// CFC twin of T_SafeConnection_Tests: the same tests drawn as CFC diagrams, the way a TwinSAFE project is authored.
    FUNCTION_BLOCK T_SafeConnection_Tests_CFC EXTENDS T_SafeCfcTestSuite
    VAR
    // Test_StartsUpToDataWhenGroupRuns
    group_1 : T_SafeGroup;
    conn_1 : T_SafeConnection(group := group_1);
    // Test_ComErrorClearedByAcknowledge
    group_2 : T_SafeGroup;
    conn_2 : T_SafeConnection(group := group_2);
END_VAR

Test_StartsUpToDataWhenGroupRuns();
Test_ComErrorClearedByAcknowledge();

METHOD PRIVATE Test_StartsUpToDataWhenGroupRuns
// note: this text did not pass the execution check against the stored diagram
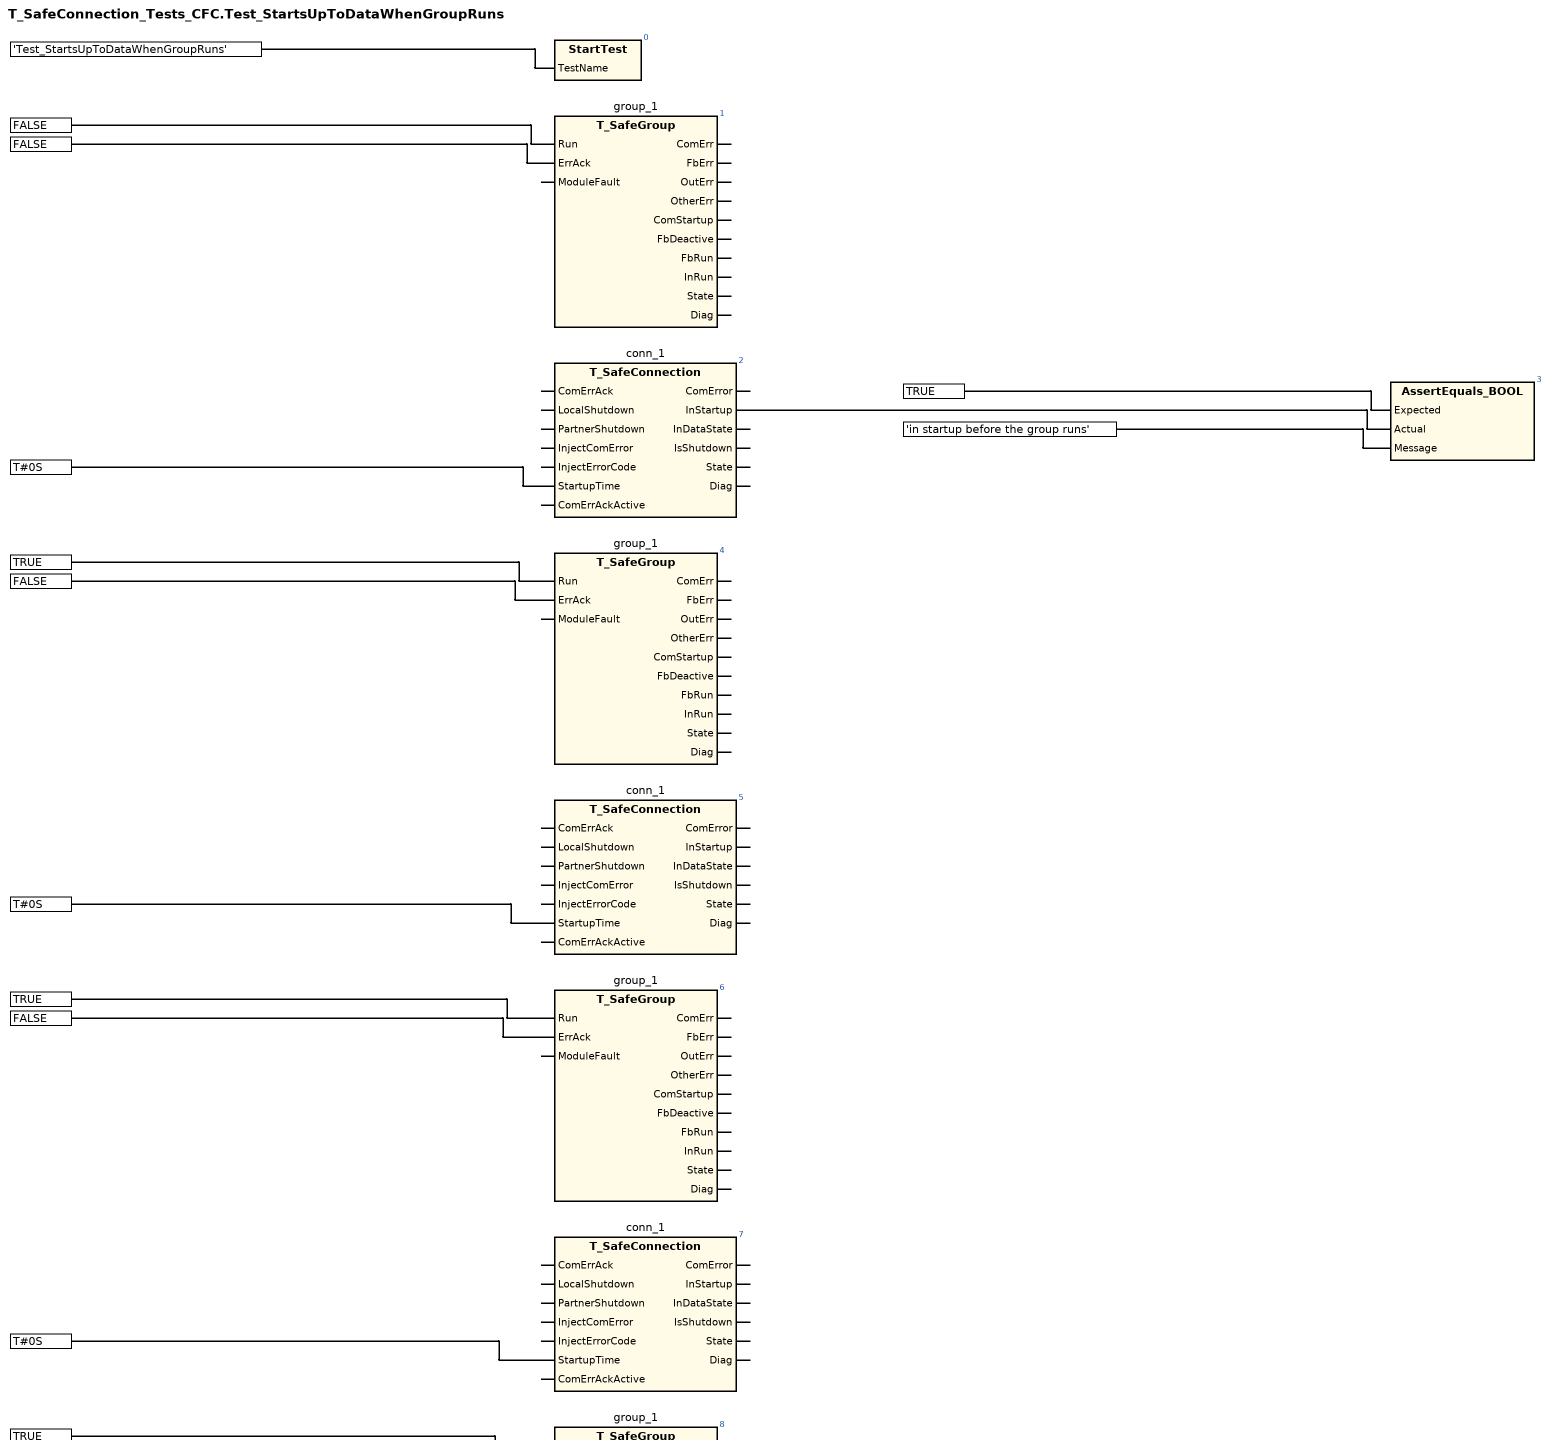
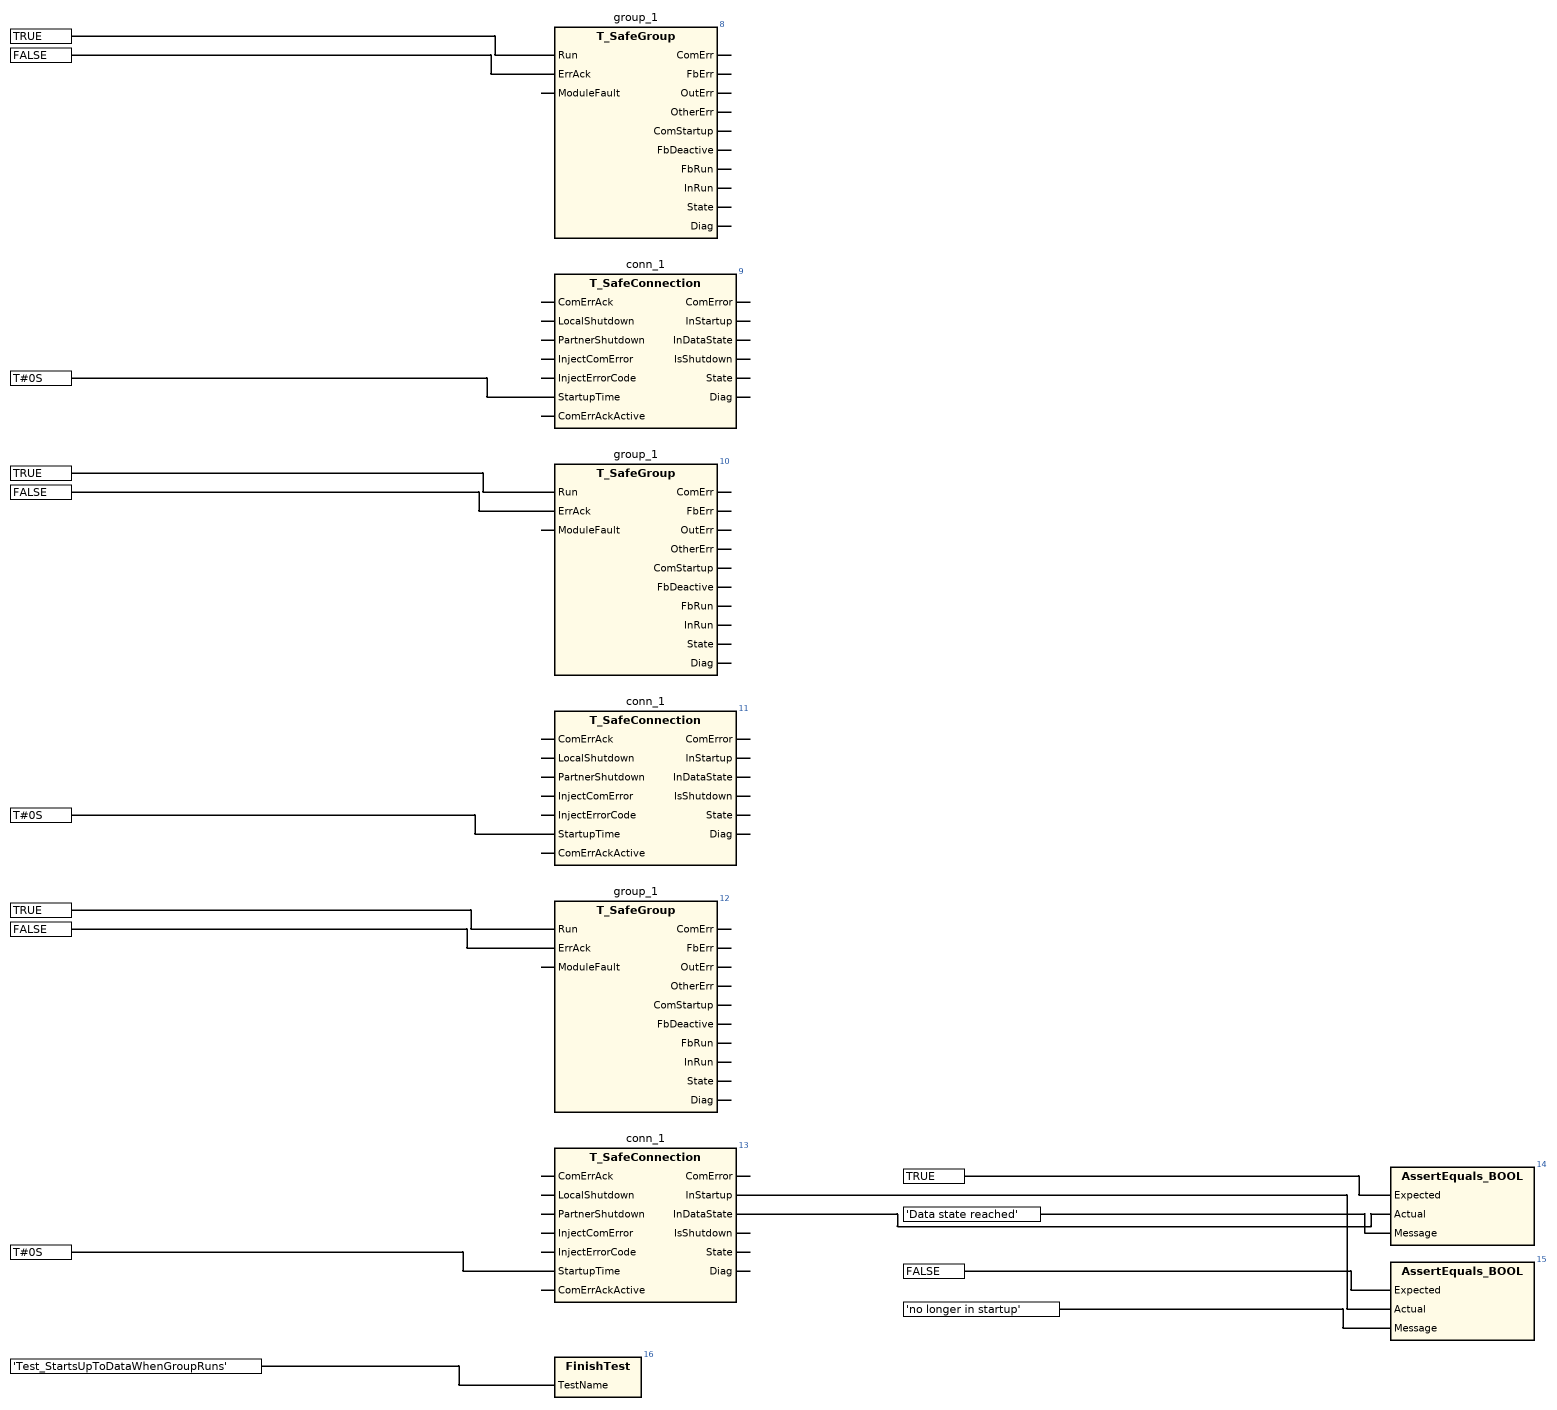
StartTest(TestName := 'Test_StartsUpToDataWhenGroupRuns');
group_1(Run := FALSE, ErrAck := FALSE); // T_SafeGroup
conn_1(StartupTime := T#0S); // T_SafeConnection
AssertEquals_BOOL(Expected := TRUE, Actual := conn_1.InStartup, Message := 'in startup before the group runs');
group_1(Run := TRUE, ErrAck := FALSE); // T_SafeGroup
conn_1(StartupTime := T#0S); // T_SafeConnection
group_1(Run := TRUE, ErrAck := FALSE); // T_SafeGroup
conn_1(StartupTime := T#0S); // T_SafeConnection
group_1(Run := TRUE, ErrAck := FALSE); // T_SafeGroup
conn_1(StartupTime := T#0S); // T_SafeConnection
group_1(Run := TRUE, ErrAck := FALSE); // T_SafeGroup
conn_1(StartupTime := T#0S); // T_SafeConnection
group_1(Run := TRUE, ErrAck := FALSE); // T_SafeGroup
conn_1(StartupTime := T#0S); // T_SafeConnection
AssertEquals_BOOL(Expected := TRUE, Actual := conn_1.InDataState, Message := 'Data state reached');
AssertEquals_BOOL(Expected := FALSE, Actual := conn_1.InStartup, Message := 'no longer in startup');
FinishTest(TestName := 'Test_StartsUpToDataWhenGroupRuns');
END_METHOD

METHOD PRIVATE Test_ComErrorClearedByAcknowledge
// note: this text did not pass the execution check against the stored diagram
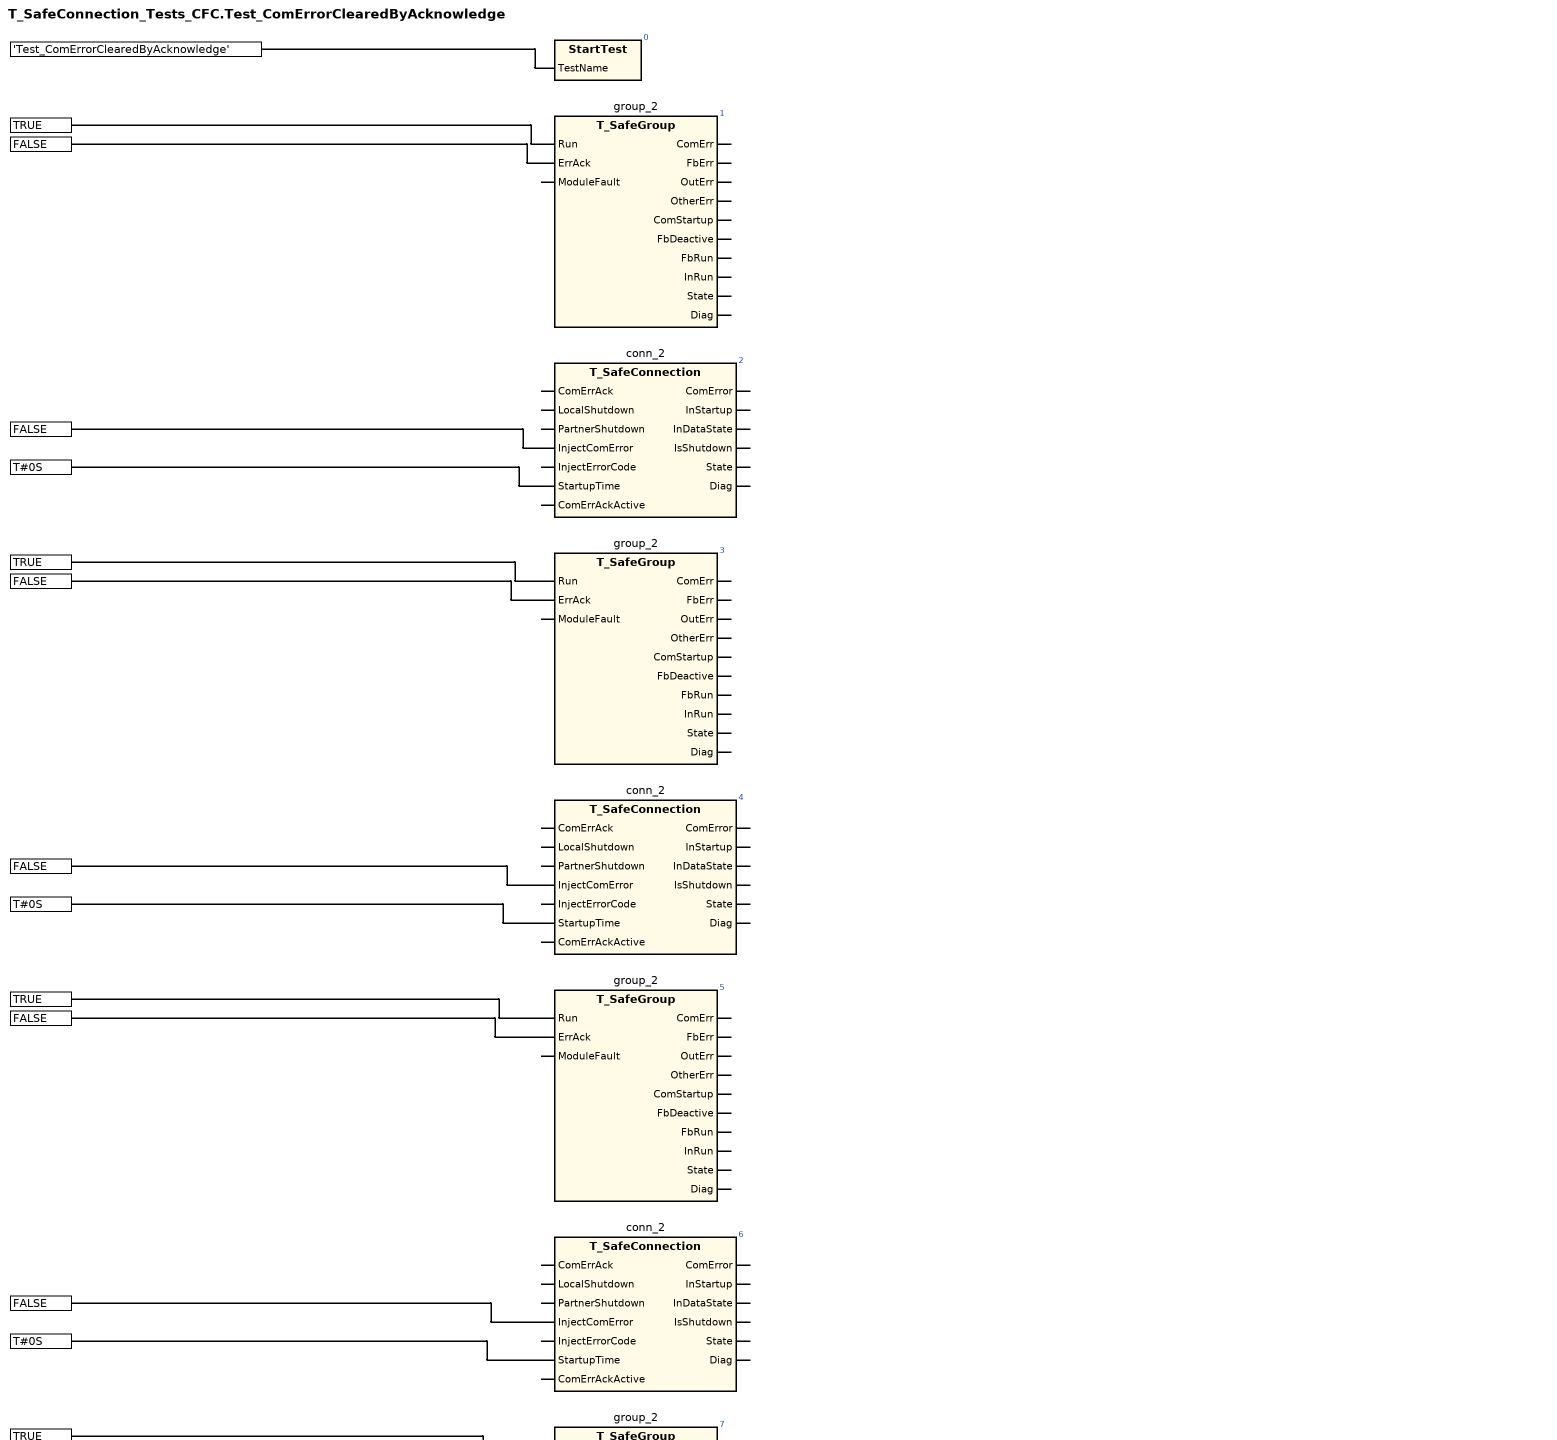
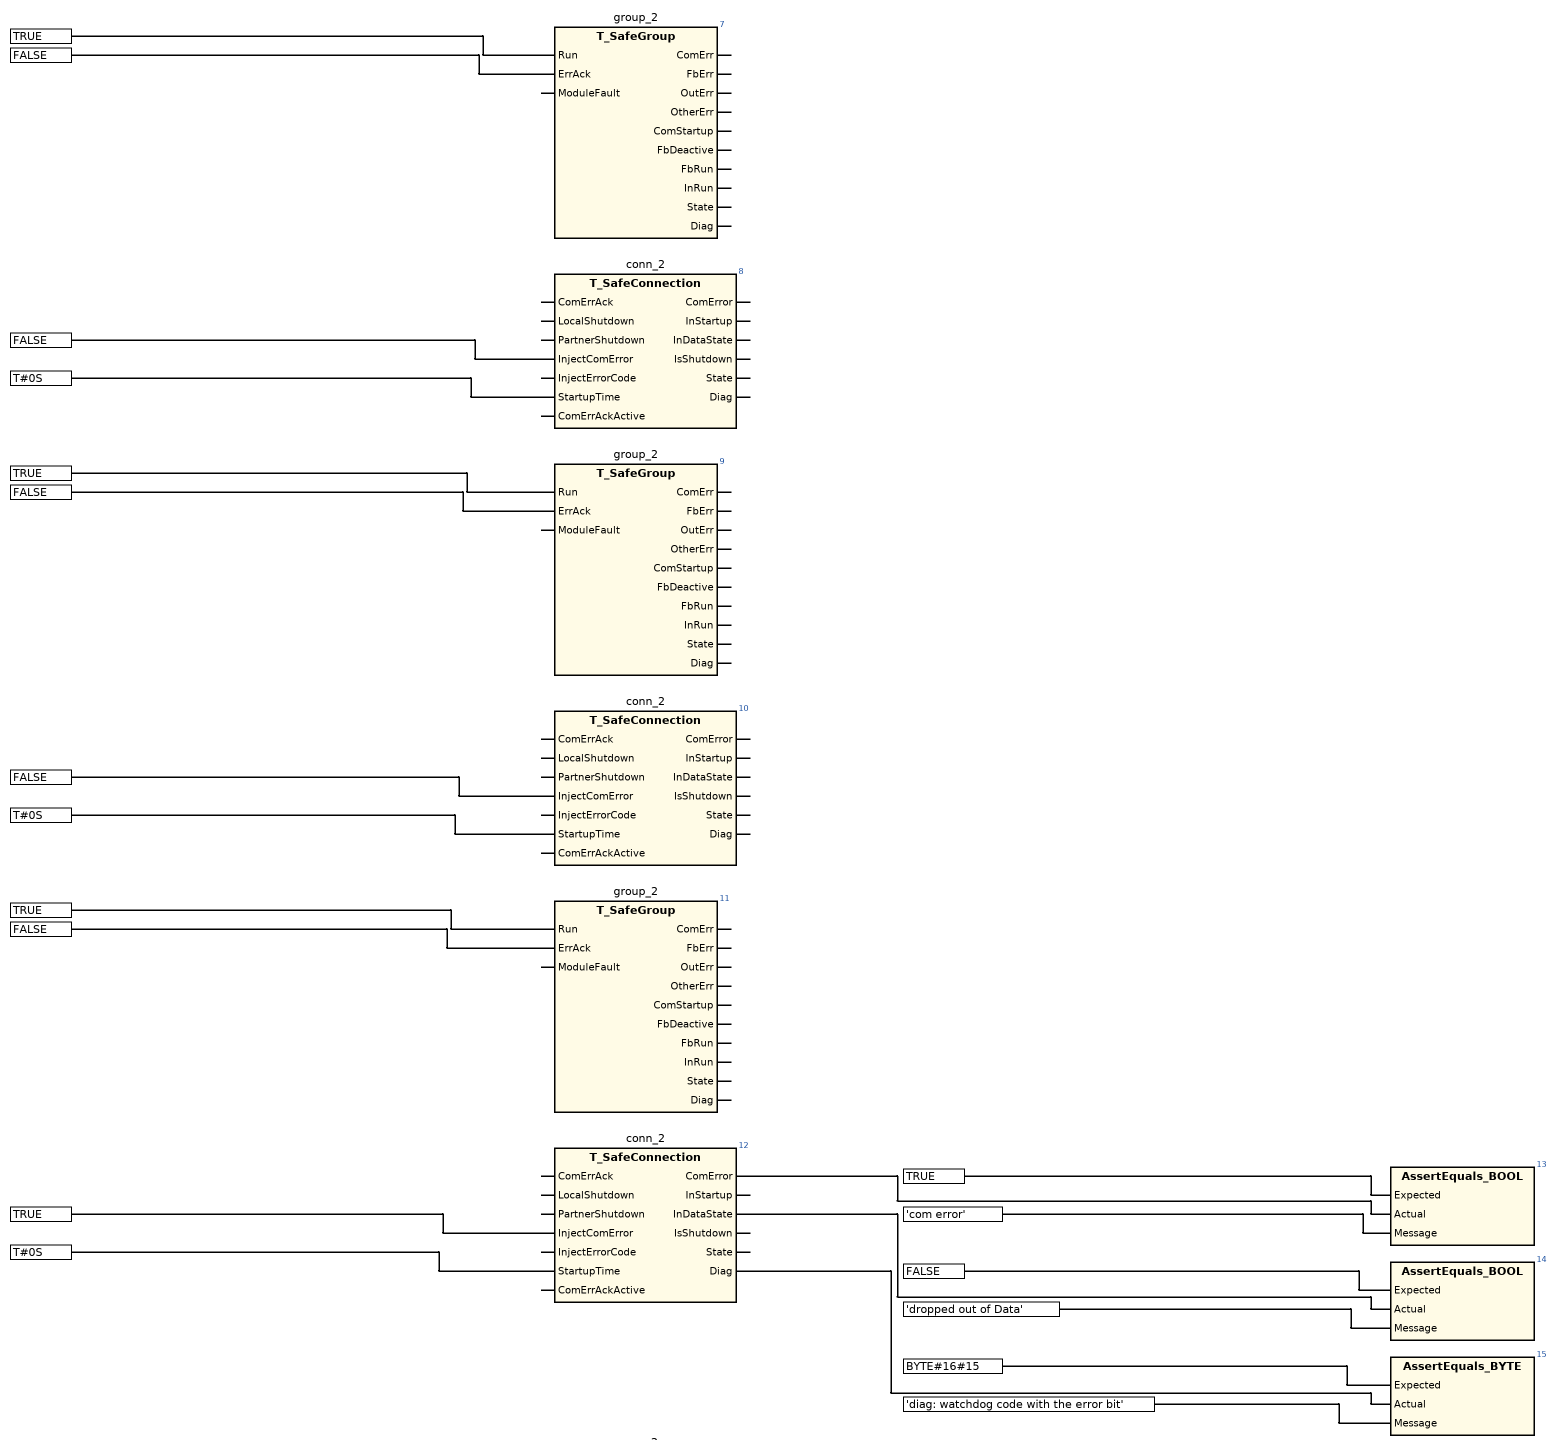
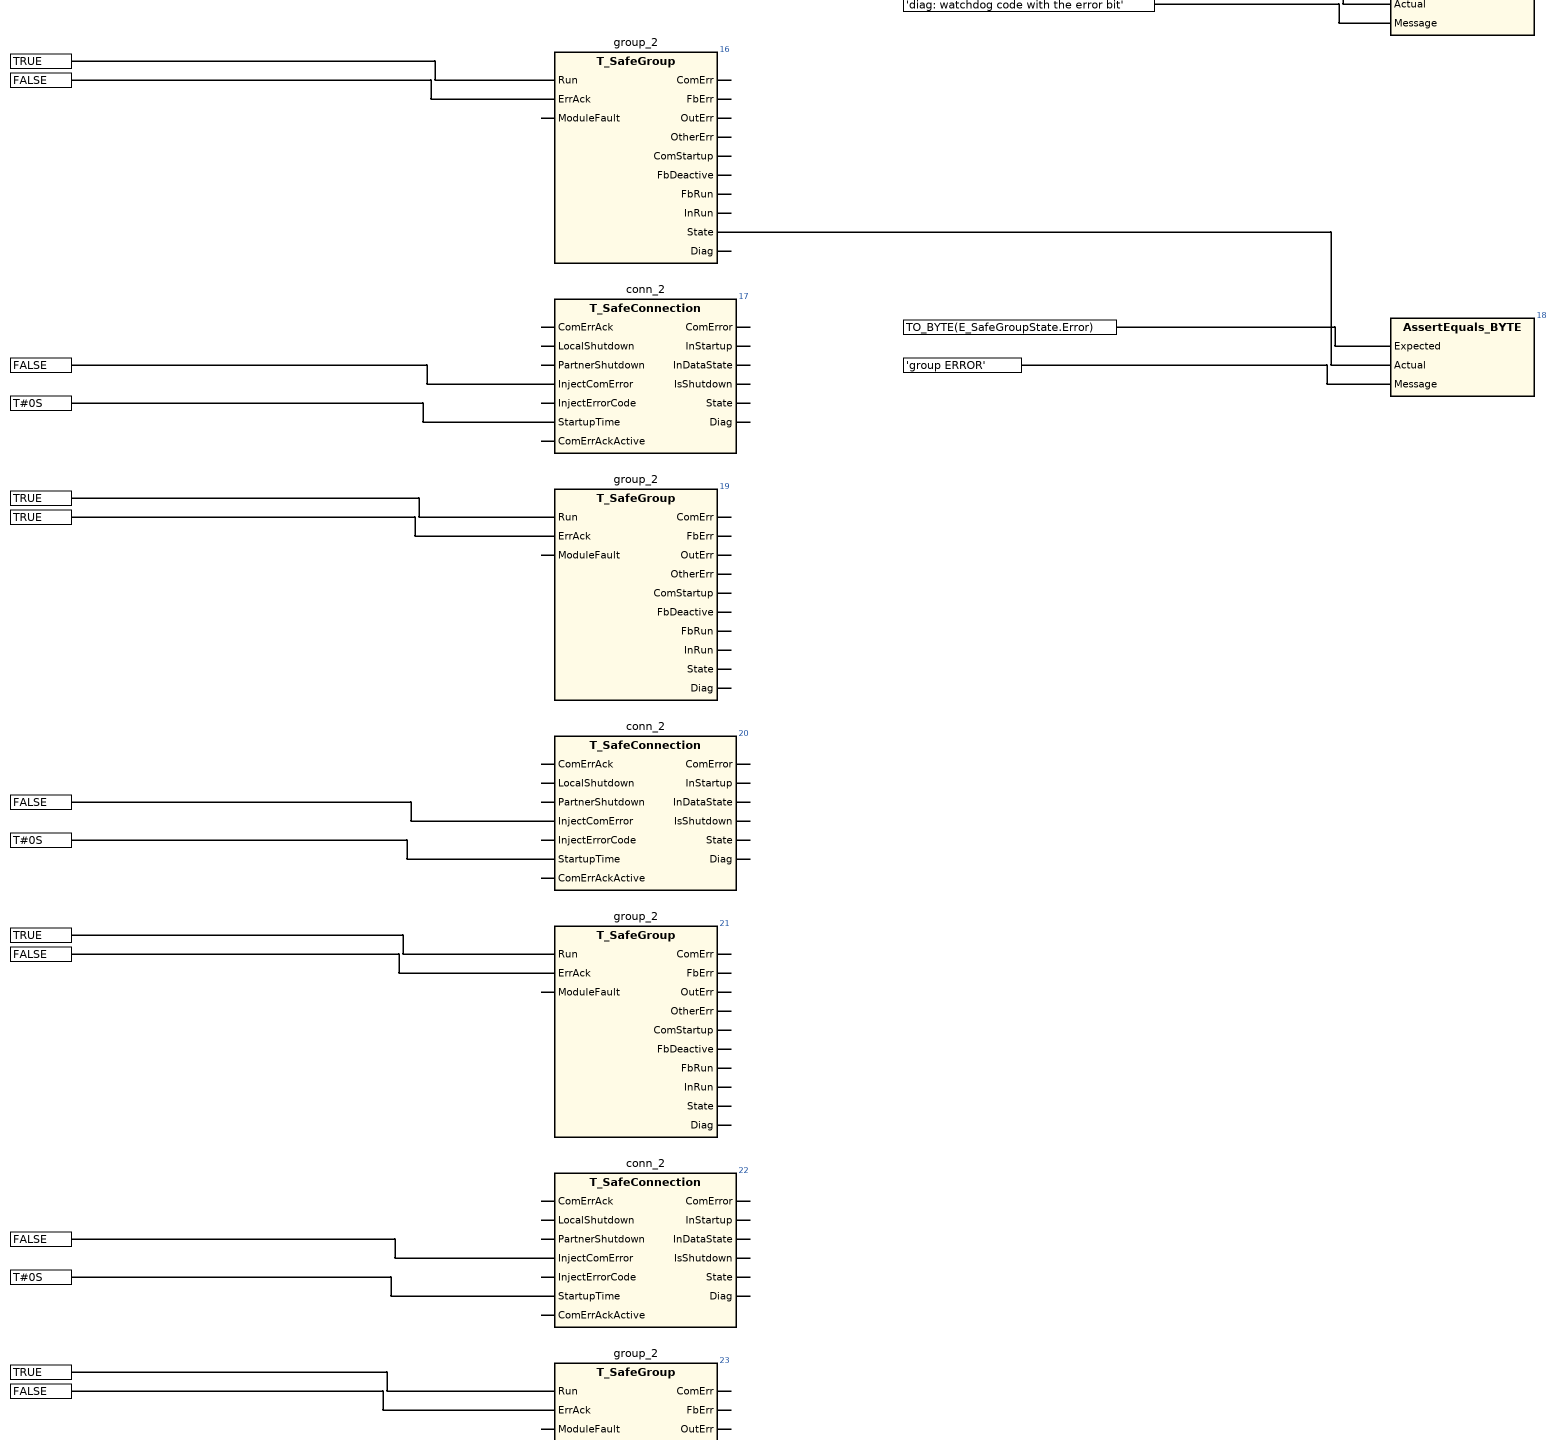
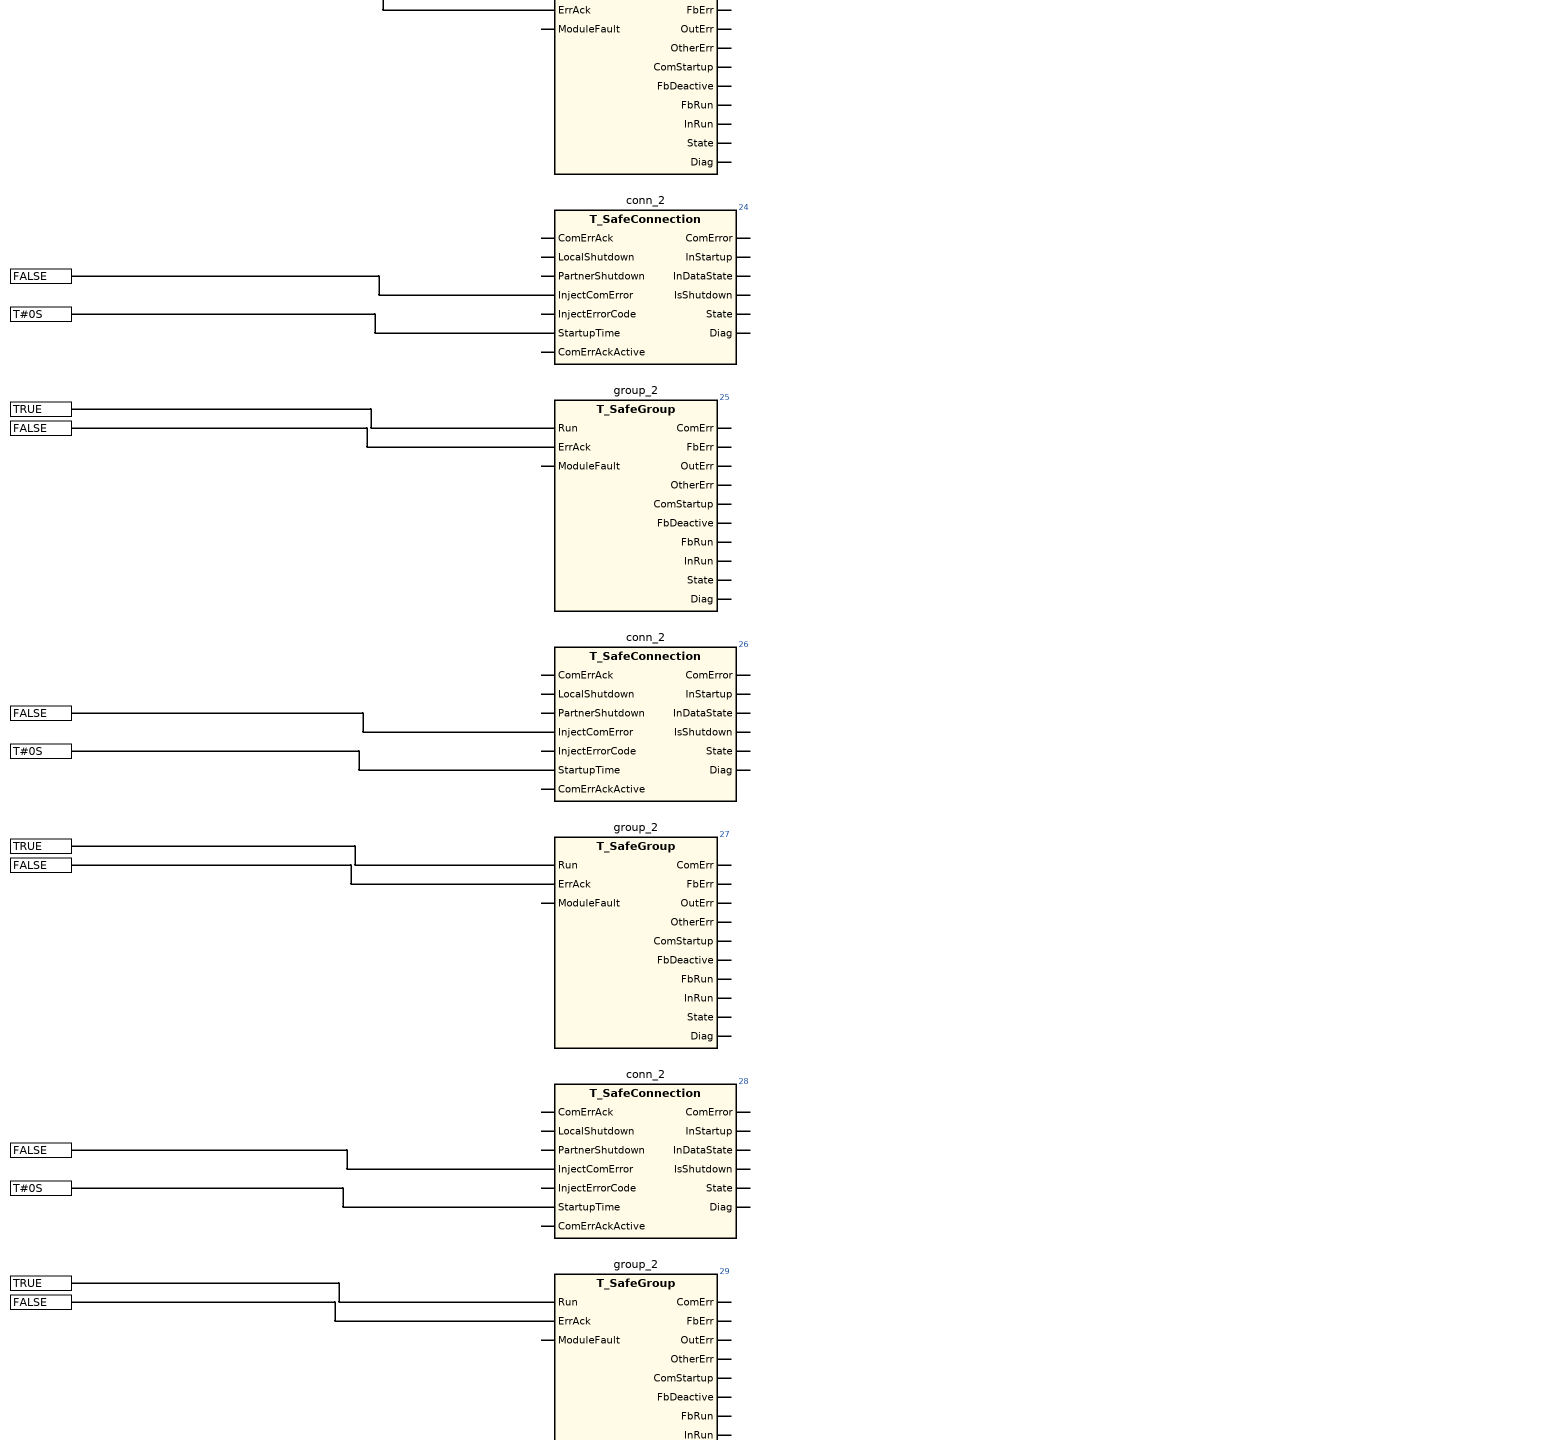
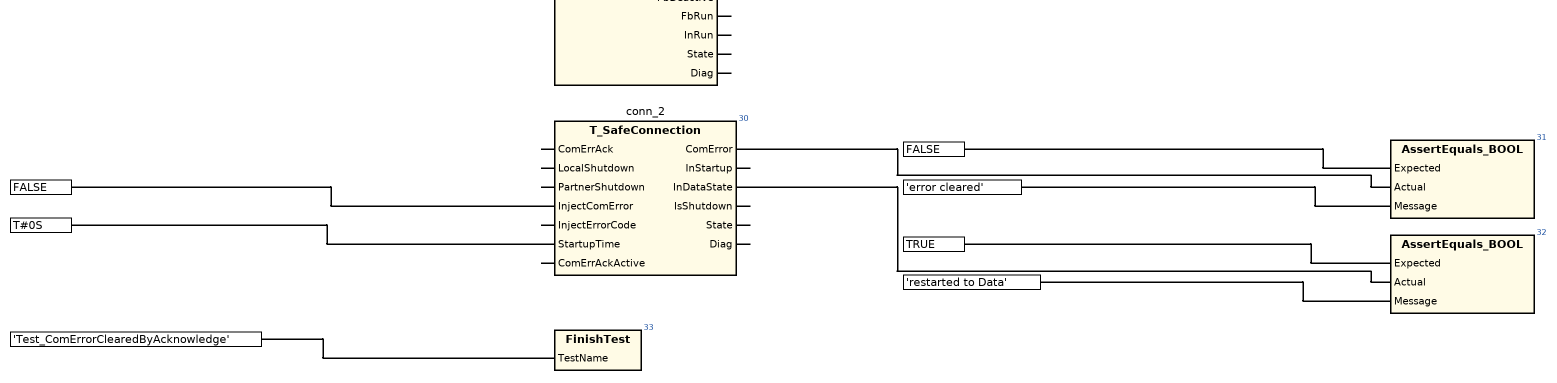
StartTest(TestName := 'Test_ComErrorClearedByAcknowledge');
group_2(Run := TRUE, ErrAck := FALSE); // T_SafeGroup
conn_2(InjectComError := FALSE, StartupTime := T#0S); // T_SafeConnection
group_2(Run := TRUE, ErrAck := FALSE); // T_SafeGroup
conn_2(InjectComError := FALSE, StartupTime := T#0S); // T_SafeConnection
group_2(Run := TRUE, ErrAck := FALSE); // T_SafeGroup
conn_2(InjectComError := FALSE, StartupTime := T#0S); // T_SafeConnection
group_2(Run := TRUE, ErrAck := FALSE); // T_SafeGroup
conn_2(InjectComError := FALSE, StartupTime := T#0S); // T_SafeConnection
group_2(Run := TRUE, ErrAck := FALSE); // T_SafeGroup
conn_2(InjectComError := FALSE, StartupTime := T#0S); // T_SafeConnection
group_2(Run := TRUE, ErrAck := FALSE); // T_SafeGroup
conn_2(InjectComError := TRUE, StartupTime := T#0S); // T_SafeConnection
AssertEquals_BOOL(Expected := TRUE, Actual := conn_2.ComError, Message := 'com error');
AssertEquals_BOOL(Expected := FALSE, Actual := conn_2.InDataState, Message := 'dropped out of Data');
AssertEquals_BYTE(Expected := BYTE#16#15, Actual := conn_2.Diag, Message := 'diag: watchdog code with the error bit');
group_2(Run := TRUE, ErrAck := FALSE); // T_SafeGroup
conn_2(InjectComError := FALSE, StartupTime := T#0S); // T_SafeConnection
AssertEquals_BYTE(Expected := TO_BYTE(E_SafeGroupState.Error), Actual := group_2.State, Message := 'group ERROR');
group_2(Run := TRUE, ErrAck := TRUE); // T_SafeGroup
conn_2(InjectComError := FALSE, StartupTime := T#0S); // T_SafeConnection
group_2(Run := TRUE, ErrAck := FALSE); // T_SafeGroup
conn_2(InjectComError := FALSE, StartupTime := T#0S); // T_SafeConnection
group_2(Run := TRUE, ErrAck := FALSE); // T_SafeGroup
conn_2(InjectComError := FALSE, StartupTime := T#0S); // T_SafeConnection
group_2(Run := TRUE, ErrAck := FALSE); // T_SafeGroup
conn_2(InjectComError := FALSE, StartupTime := T#0S); // T_SafeConnection
group_2(Run := TRUE, ErrAck := FALSE); // T_SafeGroup
conn_2(InjectComError := FALSE, StartupTime := T#0S); // T_SafeConnection
group_2(Run := TRUE, ErrAck := FALSE); // T_SafeGroup
conn_2(InjectComError := FALSE, StartupTime := T#0S); // T_SafeConnection
AssertEquals_BOOL(Expected := FALSE, Actual := conn_2.ComError, Message := 'error cleared');
AssertEquals_BOOL(Expected := TRUE, Actual := conn_2.InDataState, Message := 'restarted to Data');
FinishTest(TestName := 'Test_ComErrorClearedByAcknowledge');
END_METHOD

END_FUNCTION_BLOCK

(* stored: Version 1.1.0.1, ProductVersion 3.1.4026.22
   POU T_SafeConnection_Tests_CFC: Id {578b98aa-5be7-57b0-b00b-107f5847fc38}, SpecialFunc None
   Method Test_StartsUpToDataWhenGroupRuns: Id {bbc67d94-3fb8-528a-b4cd-99e22d8da650}
   Method Test_ComErrorClearedByAcknowledge: Id {e721ca15-6814-55e9-ba69-59e903e43b7a} *)
